(* IEC 61131-3 sources: rusty/tests/lit/single/literals, 7 files *)

(* ---- floating_point.st ---- *)
// RUN: %COMPILE %s && %RUN | %CHECK %s
VAR_GLOBAL
    // Basic global variables
    g_LREAL_pos : LREAL := 12.1212;
    g_LREAL_neg : LREAL := -12.1212;
    g_REAL_pos : REAL := 15.62;
    g_REAL_neg : REAL := -15.62;

    // Edge cases - very large numbers (should trigger LREAL inference)
    g_LREAL_huge : LREAL := 1e100;
    g_LREAL_huge_neg : LREAL := -1e100;

    // Edge cases - very small numbers (close to zero)
    g_LREAL_tiny : LREAL := 1e-100;
    g_LREAL_tiny_neg : LREAL := -1e-100;

    // High precision numbers (should preserve precision in LREAL)
    g_LREAL_precise : LREAL := 1.23456789012345678901234567890;
    g_REAL_precise : REAL := 1.23456789012345678901234567890;

    // Numbers at f32 limits
    g_LREAL_f32_max : LREAL := 3.4028235e38;
    g_LREAL_over_f32 : LREAL := 3.5e38;
END_VAR

FUNCTION main
VAR
    // Function-local variables with edge cases
    valueLREAL : LREAL := 3.14;
    valueREAL : REAL := 3.14;
    valueLREAL_neg : LREAL := -3.14159;
    valueREAL_neg : REAL := -3.14159;
    funcLREAL_huge : LREAL := 1e100;
    funcREAL_precise : REAL := 1.234567890123456789;
    funcLREAL_tiny : LREAL := 1e-200;
    funcREAL_tiny : REAL := 1e-20;
END_VAR
    // Function Local Variables
    // CHECK: Function LREAL: 3.140000
    printf('Function LREAL: %f$N', valueLREAL);
    // CHECK: Function REAL: 3.140000
    printf('Function REAL: %f$N', valueREAL);
    // CHECK: Function LREAL negative: -3.141590
    printf('Function LREAL negative: %f$N', valueLREAL_neg);
    // CHECK: Function REAL negative: -3.141590
    printf('Function REAL negative: %f$N', valueREAL_neg);

    // Function Edge Cases
    // CHECK: Function LREAL huge: 1.000000e+100
    printf('Function LREAL huge: %e$N', funcLREAL_huge);
    // CHECK: Function REAL precise: 1.234568
    printf('Function REAL precise: %f$N', funcREAL_precise);
    // CHECK: Function LREAL tiny: 1.000000e-200
    printf('Function LREAL tiny: %e$N', funcLREAL_tiny);

    // Global Variables
    // CHECK: Global LREAL positive: 12.121200
    printf('Global LREAL positive: %f$N', g_LREAL_pos);
    // CHECK: Global LREAL negative: -12.121200
    printf('Global LREAL negative: %f$N', g_LREAL_neg);
    // CHECK: Global REAL positive: 15.620000
    printf('Global REAL positive: %f$N', g_REAL_pos);
    // CHECK: Global REAL negative: -15.620000
    printf('Global REAL negative: %f$N', g_REAL_neg);

    // Global Edge Cases
    // CHECK: Global LREAL huge: 1.000000e+100
    printf('Global LREAL huge: %e$N', g_LREAL_huge);
    // CHECK: Global LREAL huge neg: -1.000000e+100
    printf('Global LREAL huge neg: %e$N', g_LREAL_huge_neg);
    // CHECK: Global LREAL tiny: 1.000000e-100
    printf('Global LREAL tiny: %e$N', g_LREAL_tiny);
    // CHECK: Global LREAL tiny neg: -1.000000e-100
    printf('Global LREAL tiny neg: %e$N', g_LREAL_tiny_neg);
    // CHECK: Global LREAL precise: 1.234567890123457
    printf('Global LREAL precise: %.15f$N', g_LREAL_precise);
    // CHECK: Global REAL precise: 1.234568
    printf('Global REAL precise: %f$N', g_REAL_precise);
    // CHECK: Global LREAL f32 max: 3.402823e+38
    printf('Global LREAL f32 max: %e$N', g_LREAL_f32_max);
    // CHECK: Global LREAL over f32: 3.500000e+38
    printf('Global LREAL over f32: %e$N', g_LREAL_over_f32);
END_FUNCTION

(* ---- integer_hex_binary.st ---- *)
// RUN: %COMPILE %s && %RUN | %CHECK %s

// NOTE: The runtime monitoring write API depends on these exact values.
// If this test fails, check whether the runtime parser needs a matching update.

FUNCTION main : DINT
VAR
    // Two's complement INT hex literals
    i_ffff      : INT  := 16#FFFF;
    i_8000      : INT  := 16#8000;
    i_7fff      : INT  := 16#7FFF;
    i_neg_ffff  : INT  := -16#FFFF;
    i_neg_000f  : INT  := -16#000F;

    // Two's complement DINT hex literals
    d_ffffffff  : DINT := 16#FFFFFFFF;
    d_80000000  : DINT := 16#80000000;

    // Two's complement INT binary literal
    i_bin_ffff  : INT  := 2#1111111111111111;
END_VAR
    // --- INT hex ---
    // CHECK: 16#FFFF as INT: -1
    printf('16#FFFF as INT: %d$N', i_ffff);
    // CHECK: 16#8000 as INT: -32768
    printf('16#8000 as INT: %d$N', i_8000);
    // CHECK: 16#7FFF as INT: 32767
    printf('16#7FFF as INT: %d$N', i_7fff);
    // CHECK: -16#FFFF as INT: 1
    printf('-16#FFFF as INT: %d$N', i_neg_ffff);
    // CHECK: -16#000F as INT: -15
    printf('-16#000F as INT: %d$N', i_neg_000f);

    // --- DINT hex ---
    // CHECK: 16#FFFFFFFF as DINT: -1
    printf('16#FFFFFFFF as DINT: %d$N', d_ffffffff);
    // CHECK: 16#80000000 as DINT: -2147483648
    printf('16#80000000 as DINT: %d$N', d_80000000);

    // --- INT binary ---
    // CHECK: 2#1111111111111111 as INT: -1
    printf('2#1111111111111111 as INT: %d$N', i_bin_ffff);
END_FUNCTION

(* ---- temporal_exact.st ---- *)
// Temporal literals are evaluated with exact integer arithmetic: no 32-bit truncation of a
// nanosecond segment, no rounding of a fraction into the next second, and the same value whether
// the literal is written in code or converted from a string at runtime.
// RUN: %COMPILE %s && %RUN | %CHECK %s

FUNCTION main : DINT
VAR
    big_ns       : LTIME := LTIME#5000000000ns;
    fraction     : LTIME := LTIME#1.5h30m;
    plus         : TIME  := T#+1s;
    digit_groups : TIME  := T#1_000ms;
    exact_max    : LTIME := LTIME#106751d23h47m16s854ms775us807ns;
    tod_fraction : LTOD  := LTOD#23:59:59.9999999999;
    dt_fraction  : DT    := DT#2024-01-01-23:59:59.9999999999;
END_VAR
    printf('big_ns=%s$N', REF(LTIME_TO_STRING(big_ns)));             // CHECK: big_ns=LTIME#5s
    printf('fraction=%s$N', REF(LTIME_TO_STRING(fraction)));         // CHECK-NEXT: fraction=LTIME#2h
    printf('plus=%s$N', REF(TIME_TO_STRING(plus)));                  // CHECK-NEXT: plus=T#1s
    printf('digit_groups=%s$N', REF(TIME_TO_STRING(digit_groups)));  // CHECK-NEXT: digit_groups=T#1s
    printf('exact_max=%s$N', REF(LTIME_TO_STRING(exact_max)));       // CHECK-NEXT: exact_max=LTIME#106751d23h47m16s854ms775us807ns
    printf('tod_fraction=%s$N', REF(LTOD_TO_STRING(tod_fraction)));  // CHECK-NEXT: tod_fraction=LTOD#23:59:59.999999999
    printf('dt_fraction=%s$N', REF(DT_TO_STRING(dt_fraction)));      // CHECK-NEXT: dt_fraction=DT#2024-01-01-23:59:59

    printf('same_as_runtime=%d$N', big_ns = STRING_TO_LTIME('LTIME#5000000000ns') AND exact_max = STRING_TO_LTIME('LTIME#106751d23h47m16s854ms775us807ns')); // CHECK-NEXT: same_as_runtime=1
END_FUNCTION

(* ---- test_floating_simple.st ---- *)
// RUN: %COMPILE %s && %RUN | %CHECK %s

FUNCTION main : DINT
    VAR
        val : LREAL := 3.14;
    END_VAR
    // CHECK: Value: 3.140000
    printf('Value: %f$N', val);
END_FUNCTION

(* ---- test_floating_inout.st ---- *)
// RUN: %COMPILE %s && %RUN | %CHECK %s

PROGRAM testProg
VAR
    val : LREAL := 3.14;
END_VAR
VAR_IN_OUT
    ioVal : LREAL := 1.0;
    ioVal1 : LREAL;
END_VAR
    // CHECK: Value: 3.140000
    printf('Value: %f$N', val);
    // CHECK: IO Value: 1.000000
    printf('IO Value: %f$N', ioVal);
    // CHECK: IO Value: 5.000000
    printf('IO Value: %f$N', ioVal1);
END_PROGRAM

FUNCTION main : DINT
    VAR
        v : LREAL := 5.0;
        u : LREAL := 5.0;
    END_VAR
    testProg(v,u);
END_FUNCTION

(* ---- test_floating_program.st ---- *)
// RUN: %COMPILE %s && %RUN | %CHECK %s

PROGRAM testProg
VAR
    val : LREAL := 3.14;
END_VAR
    // CHECK: Value: 3.140000
    printf('Value: %f$N', val);
END_PROGRAM

FUNCTION main : DINT
    testProg();
END_FUNCTION

(* ---- test_simple_inout.st ---- *)
// RUN: %COMPILE %s && %RUN | %CHECK %s

PROGRAM testProg
VAR_IN_OUT
    ioValue : LREAL := 3.14;
END_VAR
    // CHECK: Value: 3.140000
    printf('Value: %f$N', ioValue);
END_PROGRAM

FUNCTION main : DINT
    VAR
        value : LREAL := 1.0;
    END_VAR
    testProg(value);
END_FUNCTION
